// TIA Portal V20 export
// export: Created 2026-10-12T05:35:25.6965856Z, ExportSetting WithDefaults, DisplayName Totally Integrated Automation Portal, DisplayVersion V20, DisplayName TIA Portal Openness, DisplayVersion V20, DisplayName TIA Portal Teamcenter Gateway, DisplayVersion V20, DisplayName TIA Portal Version Control Interface, DisplayVersion V20, DisplayName SINAMICS Startdrive Advanced, DisplayVersion V20 SP1 Update 2, DisplayName SINAMICS Startdrive G110M, G120, G120C, G120D, G120P, G115D, DisplayVersion V20 SP1 Update 2, DisplayName SINAMICS Startdrive G130, G150, S120, S150, SINAMICS MV, G220, S200, S210, DisplayVersion V20 SP1 Update 2, DisplayName STEP 7 Professional, DisplayVersion V20, DisplayName STEP 7 Safety, DisplayVersion V20, DisplayName WinCC Basic/Comfort/Advanced, DisplayVersion V20, DisplayName WinCC Professional, DisplayVersion V20, DisplayName WinCC Unified, DisplayVersion V20
FUNCTION "FRK_ConfigRoot" : Int   // FC102, SCL
{ S7_Optimized_Access := 'TRUE' }
VERSION : 0.1
// stored: AutoNumber true, IsIECCheckEnabled false, SetENOAutomatically false, UDAEnableTagReadback false
   VAR_INPUT
      RegIndex : DInt;
   END_VAR
BEGIN

   #FRK_ConfigRoot := 0;
   CASE #RegIndex OF
       1:
           #FRK_ConfigRoot := 1;
       2:
           #FRK_ConfigRoot := 1;
       3:
           #FRK_ConfigRoot := 1;
       4:
           #FRK_ConfigRoot := 1;
       5:
           #FRK_ConfigRoot := 1;
       6:
           #FRK_ConfigRoot := 1;
       7:
           #FRK_ConfigRoot := 1;
       8:
           #FRK_ConfigRoot := 1;
       9:
           #FRK_ConfigRoot := 1;
       10:
           #FRK_ConfigRoot := 1;
       11:
           #FRK_ConfigRoot := 1;
       12:
           #FRK_ConfigRoot := 1;
       13:
           #FRK_ConfigRoot := 2;
       14:
           #FRK_ConfigRoot := 2;
       15:
           #FRK_ConfigRoot := 2;
       16:
           #FRK_ConfigRoot := 2;
       17:
           #FRK_ConfigRoot := 2;
       18:
           #FRK_ConfigRoot := 2;
       19:
           #FRK_ConfigRoot := 2;
       20:
           #FRK_ConfigRoot := 2;
       21:
           #FRK_ConfigRoot := 2;
       22:
           #FRK_ConfigRoot := 2;
       23:
           #FRK_ConfigRoot := 2;
       24:
           #FRK_ConfigRoot := 2;
       ELSE
           RETURN;
   END_CASE;
END_FUNCTION
